// TIA Portal V21 export
FUNCTION_BLOCK "PR_5by3CylModWoRdlck"   // FB178, LAD
TITLE = 5/3Cylinder Module Without Rod Lock
{ S7_Optimized_Access := 'TRUE' }
// stored: IsIECCheckEnabled true, MemoryReserve 100, SetENOAutomatically false
   VAR_INPUT
      iResetModule : Bool;   // Reset if 1
      iResetFaults : Bool;   // Reset Fault CMD
      iEnergizeAtPwrOn : Bool;   // Energize Poweron Input
      iWorkCmd : Bool;   // Cyl Work Postion CMD
      iHomeCmd : Bool;   // Cyl Home Postion CMD
      iWorkSen : Bool;   // Cyl Work Postion Input
      iHomeSen : Bool;   // Cyl Home Postion Input
      iWorkCleartoMove : Bool;   // connect work position interlock condition healthy
      iHomeCleartoMove : Bool;   // connect home position interlock condition healthy
      iWorkPositionLeftOption : Bool;   // It is the selection of the to keep work solenoid coil on after reaching work position
      iHomePositionLeftOption : Bool;   // It is the selection of the to keep home solenoid coil on after reaching home position
      iTimeoutValue : Time;   // Time Required E.g T#500MS,T#2S
      iWorkSensDebounceVal : Time;   // Time Required E.g T#500MS,T#2S
      iHomeSensDebounceVal : Time;   // Time Required E.g T#500MS,T#2S
   END_VAR
   VAR_OUTPUT
      qWorkSol : Bool;   // Cyl Work Position Sol Output
      qHomeSol : Bool;   // Cyl Home Position Sol Output
      qWorkOver : Bool;   // 1 if Cyl at Work Position
      qHomeOver : Bool;   // 1 if Cyl at Home Position
      qModError : Bool;   // Module Error
      qErrBothSensorOn : Bool;   // 1 If both WorkSen and HomeSen inputs are high at the same time.
      qErrHomeInterlock : Bool;   // 1 If homeCleartoMove is low and home command is active.
      qErrHomeSenNotLeft : Bool;   // 1 If home position sensor did not turn off within defined time
      qErrHomeTout : Bool;   // 1 If cylinder did not reach home position within defined time
      qErrWorkInterlock : Bool;   // 1 If WorkCleartoMove is low and work command is active.
      qErrWorkSenNotLeft : Bool;   // 1 If work position sensor did not turn off within defined time
      qErrWorkTout : Bool;   // 1 If cylinder did not reach work position within defined time
      qMsgWorkPosLost : Bool;   // 1 If work position achieved and lost its position without home
      qMsgHomePosLost : Bool;   // 1 If home position achieved and lost its position without work
      qMsgBothCmdOn : Bool;   // 1 if Home & work position command on same time
   END_VAR
   VAR
      sFltRstPls : Bool;   // Stat bit for positive edge of reset fault input
      sFltEdge : Bool;   // Positive edge of fault reset input
      sWorkPosMemBit : Bool;   // Stat bit for work position memory bit
      sHomePosMemBit : Bool;   // Stat bit for Home position memory bit
      sModError : Bool;   // Stat bit for Module error
      sWorkSensDebTime : Time;   // Stat bit work sensor debounce time
      sHomeSensDebTime : Time;   // Stat bit work sensor debounce time
      sTimeoutValue : Time;   // Stat bit for time out value
      sElapsedTime : Time;   // Stat bit for time elapsed
      sDlyWorkSensDeb { S7_SetPoint := 'True'} : TON_TIME;   // On Delay for Work Sensor Debounce
      sDlyHomeSensDeb { S7_SetPoint := 'True'} : TON_TIME;   // On Delay For Home Sensor Debounce
      sDlyTimeOut { S7_SetPoint := 'True'} : TON_TIME;   // On Delay Time Out timer
      sWorkSol : Bool;
      sErrWorkTout : Bool;
      sHomeSol : Bool;
      sErrHomeTout : Bool;
      sErrBothSensorOn : Bool;
      sErrWorkInterlock : Bool;
      sErrHomeInterlock : Bool;
      sErrWorkSenNotLeft : Bool;
      sErrHomeSenNotLeft : Bool;
      sMsgHomePosLost : Bool;
      sMsgWorkPosLost : Bool;
      sPosEdge : Bool;
      sPosEdge1 : Bool;
      sRegainWrkPos : Bool;
      sRegainHomePos : Bool;
      sBothCmdOn : Bool;
      sWorkPositionLeft : Bool;
      sHomePositionLeft : Bool;
   END_VAR
   VAR_TEMP   // added for the SCL form of the ladder/FBD networks
      _w1 : Bool;
      _w2 : Bool;
      _w3 : Bool;
      _w4 : Bool;
      _w5 : Bool;
   END_VAR
BEGIN

REGION Network 1: Header
   // ==============================================================================
   //  Company: Precision Automation & Robotics India Ltd. 
   // ------------------------------------------------------------------------------
   //  Item Code:SM0101022005
   //  Author/Created by: Amiya Das
   //  Reviewed/Checked by: Atul Patwardhan
   //  First Release on: 20-01-2017
   //  Latest update on:27-01-2025 
   // ------------------------------------------------------------------------------
   //  Tested with:Simulator
   //  Engineering/Editor: TIA Portal 15 & Higher
   // ------------------------------------------------------------------------------
   //  Restrictions: No
   //  Dependencies/Requirements: NA
   // ------------------------------------------------------------------------------
   //  Change Log:
   //  Ver.	Date                            Changed by                                  Details of changes
   //  0.2           20-01-2017                  Amiya Das      	              Second release version
   //  0.3           27-01-2025                 Sujeet Rote                                qMsgBothCmdOn message is added
   //  0.4           29-01-2025                  Sujeet Rote                                Work & home position left option bit
   // ------------------------------------------------------------------------------
   // Functionality: This block is used to control a simple motion with one work 
   // position output, one home position  output, one work position sensor and one 
   // home position sensor.
   // Inputs
   // iResetModule	Bool
   // iResetFaults	Bool
   // iEnergizeAtPwrOn	Bool
   // iWorkCmd	Bool
   // iHomeCmd	Bool
   // iWorkSen	Bool
   // iHomeSen	Bool
   // iWorkCleartoMove	Bool
   // iHomeCleartoMove	Bool
   // iWorkPositionLeftOption	Bool
   // iHomePositionLeftOption	Bool
   // iTimeoutValue	Time
   // iWorkSensDebounceVal	Time
   // iHomeSensDebounceVal	Time
   // 
   // Outputs
   // qWorkSol	Bool
   // qHomeSol	Bool
   // qWorkOver	Bool
   // qHomeOver	Bool
   // qErrBothSensorOn	Bool
   // qErrHomeInterlock	Bool
   // qErrHomeSenNotLeft	Bool
   // qErrHomeTout	Bool
   // qErrWorkInterlock	Bool
   // qErrWorkSenNotLeft	Bool
   // qErrWorkTout	Bool
   // qMsgWorkPosLost	Bool
   // qMsgHomePosLost	Bool
   // qMsgBothCmdOn	Bool
   // 
   // In-outs
   // NIL
   // ------------------------------------------------------------------------------
   // Errors reported:
   // 1.qErrBothSensorOn: If both WorkSen and HomeSen inputs are high at the same time.          
   // 2.qErrHomeInterlock: If homeCleartoMove is low and home command is active.
   // 3.qErrHomeSenNotLeft: If home position sensor did not turn off within defined time 
   // 4.qErrHomeTout: If cylinder did not reach home position within defined time 
   // 5.qErrWorkInterlock: If WorkCleartoMove is low and work command is active. 
   // 7.qErrWorkSenNotLeft: If work position sensor did not turn off within defined time 
   // 8.qErrWorkTout: If cylinder did not reach work position within defined time 
   // 9.qErrPipeSwaped: If Pipe or sensor swapped
   // 
   // Messages reported:
   // 1.qMsgHomePosLost: If home position achieved and lost its position without work
   // 2.qMsgWorkPosLost: If work position achieved and lost its position without home 
   // 3.qMsgBothCmdOn :  Home & work position command on same time
   // ==============================================================================
END_REGION

REGION Network 2: Fault Reset Pulse
   // Fault Reset Pulse
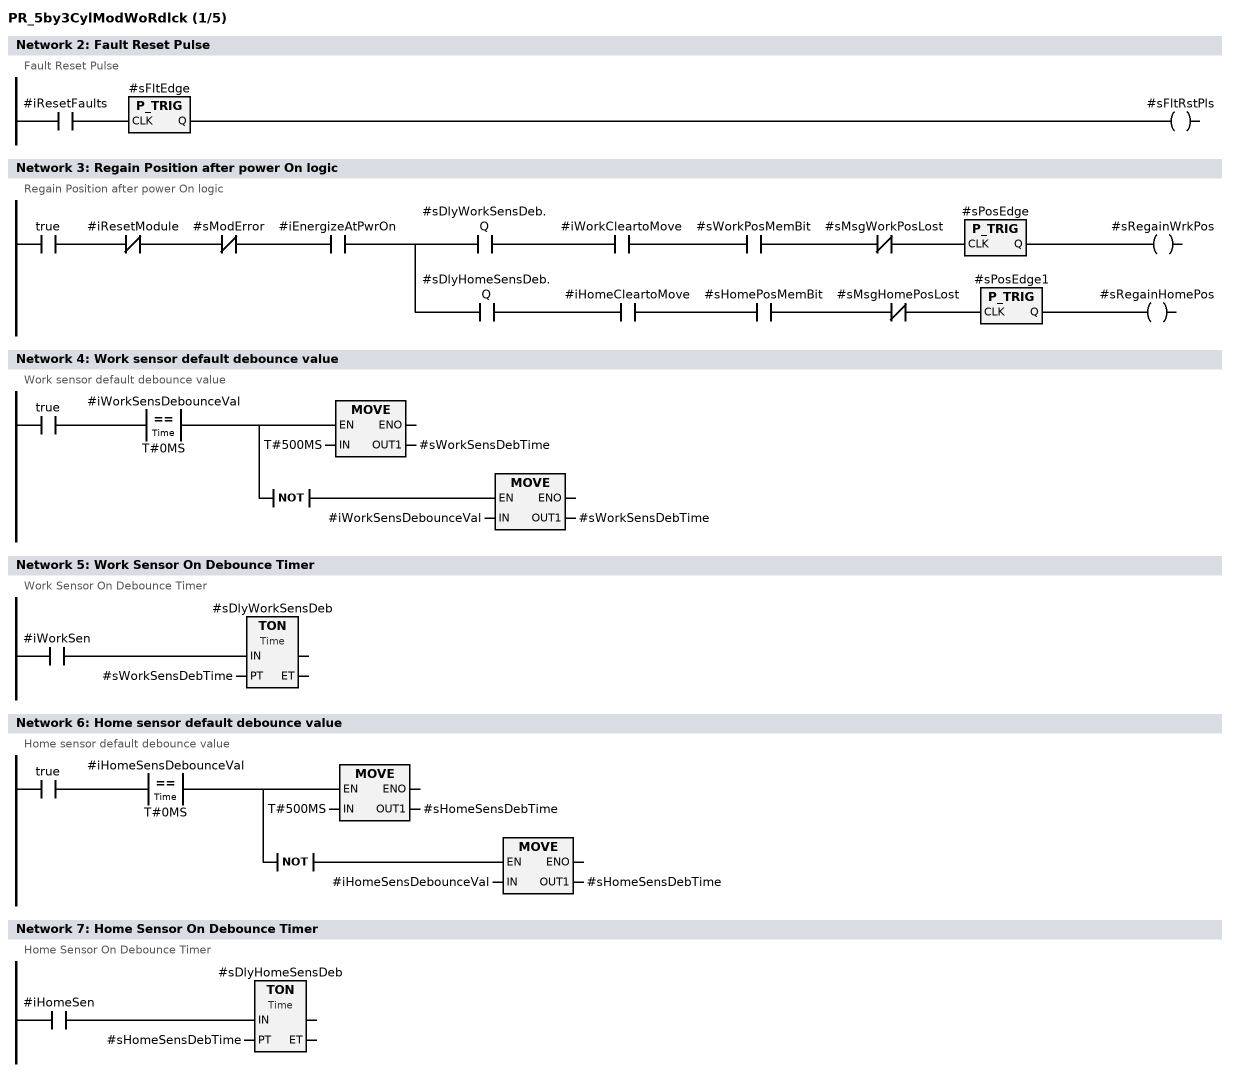
   RUNG wire#powerrail
      Contact( #iResetFaults )
      P_Trig( #sFltEdge )
      Coil( #sFltRstPls )
   END_RUNG
   // the same network as SCL:
   #_w1 := #iResetFaults AND NOT #sFltEdge;   // rising edge
   #sFltEdge := #iResetFaults;
   #sFltRstPls := #_w1;
END_REGION

REGION Network 3: Regain Position after power On logic
   // Regain Position after power On logic
   RUNG wire#powerrail
      Contact( true )
      I_Contact( #iResetModule )
      I_Contact( #sModError )
      Contact( #iEnergizeAtPwrOn )
      wire#w1
      Contact( #sDlyWorkSensDeb.Q )
      Contact( #iWorkCleartoMove )
      Contact( #sWorkPosMemBit )
      I_Contact( #sMsgWorkPosLost )
      P_Trig( #sPosEdge )
      Coil( #sRegainWrkPos )
   END_RUNG
   RUNG wire#w1
      Contact( #sDlyHomeSensDeb.Q )
      Contact( #iHomeCleartoMove )
      Contact( #sHomePosMemBit )
      I_Contact( #sMsgHomePosLost )
      P_Trig( #sPosEdge1 )
      Coil( #sRegainHomePos )
   END_RUNG
   // the same network as SCL:
   #_w1 := true AND NOT #iResetModule AND NOT #sModError AND #iEnergizeAtPwrOn;
   #_w2 := #_w1 AND #sDlyWorkSensDeb.Q AND #iWorkCleartoMove AND #sWorkPosMemBit AND NOT #sMsgWorkPosLost;
   #_w3 := #_w2 AND NOT #sPosEdge;   // rising edge
   #sPosEdge := #_w2;
   #sRegainWrkPos := #_w3;
   #_w4 := #_w1 AND #sDlyHomeSensDeb.Q AND #iHomeCleartoMove AND #sHomePosMemBit AND NOT #sMsgHomePosLost;
   #_w5 := #_w4 AND NOT #sPosEdge1;   // rising edge
   #sPosEdge1 := #_w4;
   #sRegainHomePos := #_w5;
END_REGION

REGION Network 4: Work sensor default debounce value
   // Work sensor default debounce value
   RUNG wire#powerrail
      Contact( true )
      { S7_Templates := "SrcType := Time" } EQ_Contact(in1 := #iWorkSensDebounceVal, in2 := T#0MS)
      wire#w1
      Move(in := T#500MS, out1 => #sWorkSensDebTime)
   END_RUNG
   RUNG wire#w1
      Not()
      Move(in := #iWorkSensDebounceVal, out1 => #sWorkSensDebTime)
   END_RUNG
   // the same network as SCL:
   #_w1 := true AND (#iWorkSensDebounceVal = T#0MS);
   IF #_w1 THEN #sWorkSensDebTime := T#500MS; END_IF;
   IF NOT #_w1 THEN #sWorkSensDebTime := #iWorkSensDebounceVal; END_IF;
END_REGION

REGION Network 5: Work Sensor On Debounce Timer
   // Work Sensor On Debounce Timer
   RUNG wire#powerrail
      Contact( #iWorkSen )
      { S7_Templates := "time_type := Time" } #sDlyWorkSensDeb.TON(pt := #sWorkSensDebTime, et =>)
   END_RUNG
   // the same network as SCL:
   #sDlyWorkSensDeb(IN := #iWorkSen, PT := #sWorkSensDebTime);   // TON
END_REGION

REGION Network 6: Home sensor default debounce value
   // Home sensor default debounce value
   RUNG wire#powerrail
      Contact( true )
      { S7_Templates := "SrcType := Time" } EQ_Contact(in1 := #iHomeSensDebounceVal, in2 := T#0MS)
      wire#w1
      Move(in := T#500MS, out1 => #sHomeSensDebTime)
   END_RUNG
   RUNG wire#w1
      Not()
      Move(in := #iHomeSensDebounceVal, out1 => #sHomeSensDebTime)
   END_RUNG
   // the same network as SCL:
   #_w1 := true AND (#iHomeSensDebounceVal = T#0MS);
   IF #_w1 THEN #sHomeSensDebTime := T#500MS; END_IF;
   IF NOT #_w1 THEN #sHomeSensDebTime := #iHomeSensDebounceVal; END_IF;
END_REGION

REGION Network 7: Home Sensor On Debounce Timer
   // Home Sensor On Debounce Timer
   RUNG wire#powerrail
      Contact( #iHomeSen )
      { S7_Templates := "time_type := Time" } #sDlyHomeSensDeb.TON(pt := #sHomeSensDebTime, et =>)
   END_RUNG
   // the same network as SCL:
   #sDlyHomeSensDeb(IN := #iHomeSen, PT := #sHomeSensDebTime);   // TON
END_REGION

REGION Network 8: Timeout Value
   // Timeout Value
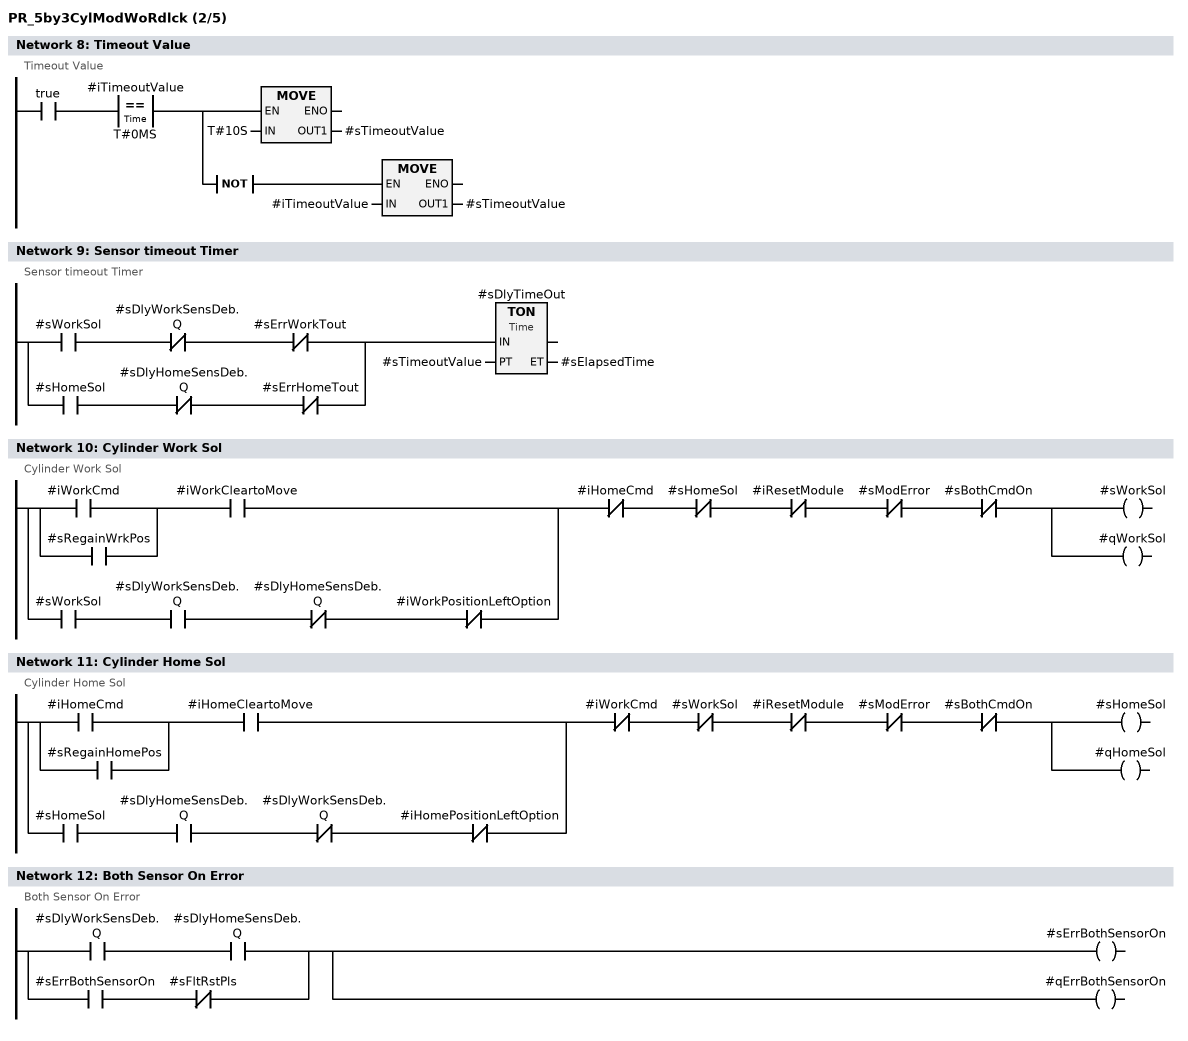
   RUNG wire#powerrail
      Contact( true )
      { S7_Templates := "SrcType := Time" } EQ_Contact(in1 := #iTimeoutValue, in2 := T#0MS)
      wire#w1
      Move(in := T#10S, out1 => #sTimeoutValue)
   END_RUNG
   RUNG wire#w1
      Not()
      Move(in := #iTimeoutValue, out1 => #sTimeoutValue)
   END_RUNG
   // the same network as SCL:
   #_w1 := true AND (#iTimeoutValue = T#0MS);
   IF #_w1 THEN #sTimeoutValue := T#10S; END_IF;
   IF NOT #_w1 THEN #sTimeoutValue := #iTimeoutValue; END_IF;
END_REGION

REGION Network 9: Sensor timeout Timer
   // Sensor timeout Timer
   RUNG wire#powerrail
      Contact( #sWorkSol )
      I_Contact( #sDlyWorkSensDeb.Q )
      I_Contact( #sErrWorkTout )
      wire#w1
      { S7_Templates := "time_type := Time" } #sDlyTimeOut.TON(pt := #sTimeoutValue, et => #sElapsedTime)
   END_RUNG
   RUNG wire#powerrail
      Contact( #sHomeSol )
      I_Contact( #sDlyHomeSensDeb.Q )
      I_Contact( #sErrHomeTout )
   END_RUNG wire#w1
   // the same network as SCL:
   #sDlyTimeOut(IN := (#sWorkSol AND NOT #sDlyWorkSensDeb.Q AND NOT #sErrWorkTout) OR (#sHomeSol AND NOT #sDlyHomeSensDeb.Q AND NOT #sErrHomeTout),   // TON
                PT := #sTimeoutValue,
                ET => #sElapsedTime);
END_REGION

REGION Network 10: Cylinder Work Sol
   // Cylinder Work Sol
   RUNG wire#powerrail
      Contact( #iWorkCmd )
      wire#w1
      Contact( #iWorkCleartoMove )
      wire#w2
      I_Contact( #iHomeCmd )
      I_Contact( #sHomeSol )
      I_Contact( #iResetModule )
      I_Contact( #sModError )
      I_Contact( #sBothCmdOn )
      wire#w3
      Coil( #sWorkSol )
   END_RUNG
   RUNG wire#powerrail
      Contact( #sRegainWrkPos )
   END_RUNG wire#w1
   RUNG wire#powerrail
      Contact( #sWorkSol )
      Contact( #sDlyWorkSensDeb.Q )
      I_Contact( #sDlyHomeSensDeb.Q )
      I_Contact( #iWorkPositionLeftOption )
   END_RUNG wire#w2
   RUNG wire#w3
      Coil( #qWorkSol )
   END_RUNG
   // the same network as SCL:
   #sWorkSol := (((#iWorkCmd OR #sRegainWrkPos) AND #iWorkCleartoMove) OR (#sWorkSol AND #sDlyWorkSensDeb.Q AND NOT #sDlyHomeSensDeb.Q AND NOT #iWorkPositionLeftOption)) AND NOT #iHomeCmd AND NOT #sHomeSol AND NOT #iResetModule AND NOT #sModError AND NOT #sBothCmdOn;
   #qWorkSol := #sWorkSol;
END_REGION

REGION Network 11: Cylinder Home Sol
   // Cylinder Home Sol
   RUNG wire#powerrail
      Contact( #iHomeCmd )
      wire#w1
      Contact( #iHomeCleartoMove )
      wire#w2
      I_Contact( #iWorkCmd )
      I_Contact( #sWorkSol )
      I_Contact( #iResetModule )
      I_Contact( #sModError )
      I_Contact( #sBothCmdOn )
      wire#w3
      Coil( #sHomeSol )
   END_RUNG
   RUNG wire#powerrail
      Contact( #sRegainHomePos )
   END_RUNG wire#w1
   RUNG wire#powerrail
      Contact( #sHomeSol )
      Contact( #sDlyHomeSensDeb.Q )
      I_Contact( #sDlyWorkSensDeb.Q )
      I_Contact( #iHomePositionLeftOption )
   END_RUNG wire#w2
   RUNG wire#w3
      Coil( #qHomeSol )
   END_RUNG
   // the same network as SCL:
   #sHomeSol := (((#iHomeCmd OR #sRegainHomePos) AND #iHomeCleartoMove) OR (#sHomeSol AND #sDlyHomeSensDeb.Q AND NOT #sDlyWorkSensDeb.Q AND NOT #iHomePositionLeftOption)) AND NOT #iWorkCmd AND NOT #sWorkSol AND NOT #iResetModule AND NOT #sModError AND NOT #sBothCmdOn;
   #qHomeSol := #sHomeSol;
END_REGION

REGION Network 12: Both Sensor On Error
   // Both Sensor On Error
   RUNG wire#powerrail
      Contact( #sDlyWorkSensDeb.Q )
      Contact( #sDlyHomeSensDeb.Q )
      wire#w1
      Coil( #sErrBothSensorOn )
   END_RUNG
   RUNG wire#powerrail
      Contact( #sErrBothSensorOn )
      I_Contact( #sFltRstPls )
   END_RUNG wire#w1
   RUNG wire#w1
      Coil( #qErrBothSensorOn )
   END_RUNG
   // the same network as SCL:
   #sErrBothSensorOn := (#sDlyWorkSensDeb.Q AND #sDlyHomeSensDeb.Q) OR (#sErrBothSensorOn AND NOT #sFltRstPls);
   #qErrBothSensorOn := #sErrBothSensorOn;
END_REGION

REGION Network 13: Work Interlock Error
   // Work Interlock Error
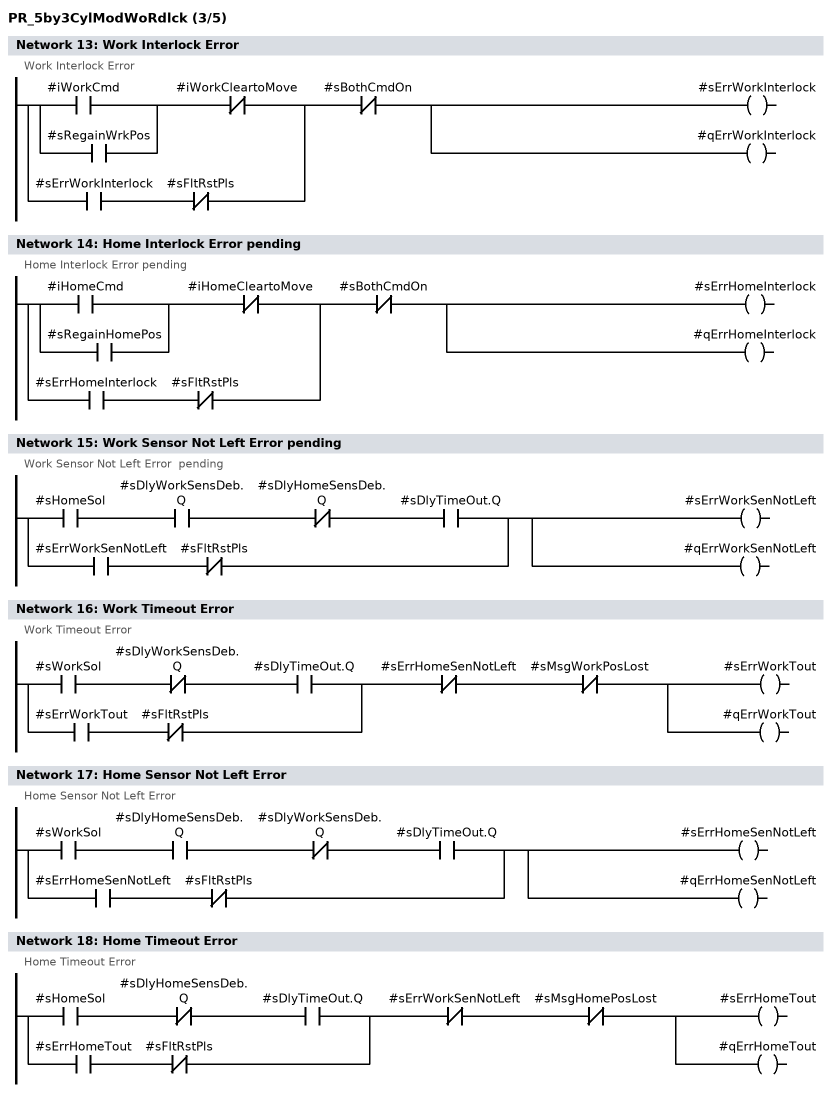
   RUNG wire#powerrail
      Contact( #iWorkCmd )
      wire#w1
      I_Contact( #iWorkCleartoMove )
      wire#w2
      I_Contact( #sBothCmdOn )
      wire#w3
      Coil( #sErrWorkInterlock )
   END_RUNG
   RUNG wire#powerrail
      Contact( #sRegainWrkPos )
   END_RUNG wire#w1
   RUNG wire#powerrail
      Contact( #sErrWorkInterlock )
      I_Contact( #sFltRstPls )
   END_RUNG wire#w2
   RUNG wire#w3
      Coil( #qErrWorkInterlock )
   END_RUNG
   // the same network as SCL:
   #sErrWorkInterlock := (((#iWorkCmd OR #sRegainWrkPos) AND NOT #iWorkCleartoMove) OR (#sErrWorkInterlock AND NOT #sFltRstPls)) AND NOT #sBothCmdOn;
   #qErrWorkInterlock := #sErrWorkInterlock;
END_REGION

REGION Network 14: Home Interlock Error pending
   // Home Interlock Error pending
   RUNG wire#powerrail
      Contact( #iHomeCmd )
      wire#w1
      I_Contact( #iHomeCleartoMove )
      wire#w2
      I_Contact( #sBothCmdOn )
      wire#w3
      Coil( #sErrHomeInterlock )
   END_RUNG
   RUNG wire#powerrail
      Contact( #sRegainHomePos )
   END_RUNG wire#w1
   RUNG wire#powerrail
      Contact( #sErrHomeInterlock )
      I_Contact( #sFltRstPls )
   END_RUNG wire#w2
   RUNG wire#w3
      Coil( #qErrHomeInterlock )
   END_RUNG
   // the same network as SCL:
   #sErrHomeInterlock := (((#iHomeCmd OR #sRegainHomePos) AND NOT #iHomeCleartoMove) OR (#sErrHomeInterlock AND NOT #sFltRstPls)) AND NOT #sBothCmdOn;
   #qErrHomeInterlock := #sErrHomeInterlock;
END_REGION

REGION Network 15: Work Sensor Not Left Error pending
   // Work Sensor Not Left Error  pending
   RUNG wire#powerrail
      Contact( #sHomeSol )
      Contact( #sDlyWorkSensDeb.Q )
      I_Contact( #sDlyHomeSensDeb.Q )
      Contact( #sDlyTimeOut.Q )
      wire#w1
      Coil( #sErrWorkSenNotLeft )
   END_RUNG
   RUNG wire#powerrail
      Contact( #sErrWorkSenNotLeft )
      I_Contact( #sFltRstPls )
   END_RUNG wire#w1
   RUNG wire#w1
      Coil( #qErrWorkSenNotLeft )
   END_RUNG
   // the same network as SCL:
   #sErrWorkSenNotLeft := (#sHomeSol AND #sDlyWorkSensDeb.Q AND NOT #sDlyHomeSensDeb.Q AND #sDlyTimeOut.Q) OR (#sErrWorkSenNotLeft AND NOT #sFltRstPls);
   #qErrWorkSenNotLeft := #sErrWorkSenNotLeft;
END_REGION

REGION Network 16: Work Timeout Error
   // Work Timeout Error
   RUNG wire#powerrail
      Contact( #sWorkSol )
      I_Contact( #sDlyWorkSensDeb.Q )
      Contact( #sDlyTimeOut.Q )
      wire#w1
      I_Contact( #sErrHomeSenNotLeft )
      I_Contact( #sMsgWorkPosLost )
      wire#w2
      Coil( #sErrWorkTout )
   END_RUNG
   RUNG wire#powerrail
      Contact( #sErrWorkTout )
      I_Contact( #sFltRstPls )
   END_RUNG wire#w1
   RUNG wire#w2
      Coil( #qErrWorkTout )
   END_RUNG
   // the same network as SCL:
   #sErrWorkTout := ((#sWorkSol AND NOT #sDlyWorkSensDeb.Q AND #sDlyTimeOut.Q) OR (#sErrWorkTout AND NOT #sFltRstPls)) AND NOT #sErrHomeSenNotLeft AND NOT #sMsgWorkPosLost;
   #qErrWorkTout := #sErrWorkTout;
END_REGION

REGION Network 17: Home Sensor Not Left Error
   // Home Sensor Not Left Error
   RUNG wire#powerrail
      Contact( #sWorkSol )
      Contact( #sDlyHomeSensDeb.Q )
      I_Contact( #sDlyWorkSensDeb.Q )
      Contact( #sDlyTimeOut.Q )
      wire#w1
      Coil( #sErrHomeSenNotLeft )
   END_RUNG
   RUNG wire#powerrail
      Contact( #sErrHomeSenNotLeft )
      I_Contact( #sFltRstPls )
   END_RUNG wire#w1
   RUNG wire#w1
      Coil( #qErrHomeSenNotLeft )
   END_RUNG
   // the same network as SCL:
   #sErrHomeSenNotLeft := (#sWorkSol AND #sDlyHomeSensDeb.Q AND NOT #sDlyWorkSensDeb.Q AND #sDlyTimeOut.Q) OR (#sErrHomeSenNotLeft AND NOT #sFltRstPls);
   #qErrHomeSenNotLeft := #sErrHomeSenNotLeft;
END_REGION

REGION Network 18: Home Timeout Error
   // Home Timeout Error
   RUNG wire#powerrail
      Contact( #sHomeSol )
      I_Contact( #sDlyHomeSensDeb.Q )
      Contact( #sDlyTimeOut.Q )
      wire#w1
      I_Contact( #sErrWorkSenNotLeft )
      I_Contact( #sMsgHomePosLost )
      wire#w2
      Coil( #sErrHomeTout )
   END_RUNG
   RUNG wire#powerrail
      Contact( #sErrHomeTout )
      I_Contact( #sFltRstPls )
   END_RUNG wire#w1
   RUNG wire#w2
      Coil( #qErrHomeTout )
   END_RUNG
   // the same network as SCL:
   #sErrHomeTout := ((#sHomeSol AND NOT #sDlyHomeSensDeb.Q AND #sDlyTimeOut.Q) OR (#sErrHomeTout AND NOT #sFltRstPls)) AND NOT #sErrWorkSenNotLeft AND NOT #sMsgHomePosLost;
   #qErrHomeTout := #sErrHomeTout;
END_REGION

REGION Network 19: Work Position Left Stat logic / Work Position Left option bit Logic
   // Work Position Left Stat logic / Work Position Left option bit Logic
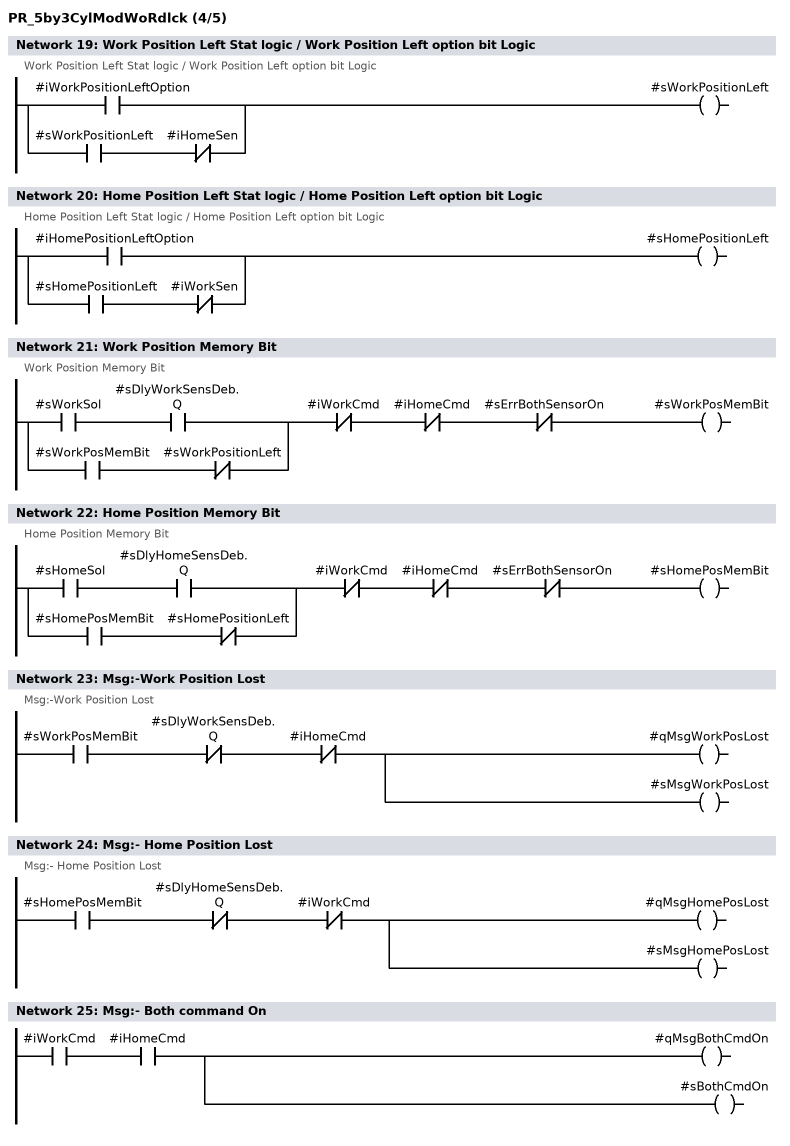
   RUNG wire#powerrail
      Contact( #iWorkPositionLeftOption )
      wire#w1
      Coil( #sWorkPositionLeft )
   END_RUNG
   RUNG wire#powerrail
      Contact( #sWorkPositionLeft )
      I_Contact( #iHomeSen )
   END_RUNG wire#w1
   // the same network as SCL:
   #sWorkPositionLeft := #iWorkPositionLeftOption OR (#sWorkPositionLeft AND NOT #iHomeSen);
END_REGION

REGION Network 20: Home Position Left Stat logic / Home Position Left option bit Logic
   // Home Position Left Stat logic / Home Position Left option bit Logic
   RUNG wire#powerrail
      Contact( #iHomePositionLeftOption )
      wire#w1
      Coil( #sHomePositionLeft )
   END_RUNG
   RUNG wire#powerrail
      Contact( #sHomePositionLeft )
      I_Contact( #iWorkSen )
   END_RUNG wire#w1
   // the same network as SCL:
   #sHomePositionLeft := #iHomePositionLeftOption OR (#sHomePositionLeft AND NOT #iWorkSen);
END_REGION

REGION Network 21: Work Position Memory Bit
   // Work Position Memory Bit
   RUNG wire#powerrail
      Contact( #sWorkSol )
      Contact( #sDlyWorkSensDeb.Q )
      wire#w1
      I_Contact( #iWorkCmd )
      I_Contact( #iHomeCmd )
      I_Contact( #sErrBothSensorOn )
      Coil( #sWorkPosMemBit )
   END_RUNG
   RUNG wire#powerrail
      Contact( #sWorkPosMemBit )
      I_Contact( #sWorkPositionLeft )
   END_RUNG wire#w1
   // the same network as SCL:
   #sWorkPosMemBit := ((#sWorkSol AND #sDlyWorkSensDeb.Q) OR (#sWorkPosMemBit AND NOT #sWorkPositionLeft)) AND NOT #iWorkCmd AND NOT #iHomeCmd AND NOT #sErrBothSensorOn;
END_REGION

REGION Network 22: Home Position Memory Bit
   // Home Position Memory Bit
   RUNG wire#powerrail
      Contact( #sHomeSol )
      Contact( #sDlyHomeSensDeb.Q )
      wire#w1
      I_Contact( #iWorkCmd )
      I_Contact( #iHomeCmd )
      I_Contact( #sErrBothSensorOn )
      Coil( #sHomePosMemBit )
   END_RUNG
   RUNG wire#powerrail
      Contact( #sHomePosMemBit )
      I_Contact( #sHomePositionLeft )
   END_RUNG wire#w1
   // the same network as SCL:
   #sHomePosMemBit := ((#sHomeSol AND #sDlyHomeSensDeb.Q) OR (#sHomePosMemBit AND NOT #sHomePositionLeft)) AND NOT #iWorkCmd AND NOT #iHomeCmd AND NOT #sErrBothSensorOn;
END_REGION

REGION Network 23: Msg:-Work Position Lost
   // Msg:-Work Position Lost
   RUNG wire#powerrail
      Contact( #sWorkPosMemBit )
      I_Contact( #sDlyWorkSensDeb.Q )
      I_Contact( #iHomeCmd )
      wire#w1
      Coil( #qMsgWorkPosLost )
   END_RUNG
   RUNG wire#w1
      Coil( #sMsgWorkPosLost )
   END_RUNG
   // the same network as SCL:
   #qMsgWorkPosLost := #sWorkPosMemBit AND NOT #sDlyWorkSensDeb.Q AND NOT #iHomeCmd;
   #sMsgWorkPosLost := #qMsgWorkPosLost;
END_REGION

REGION Network 24: Msg:- Home Position Lost
   // Msg:- Home Position Lost
   RUNG wire#powerrail
      Contact( #sHomePosMemBit )
      I_Contact( #sDlyHomeSensDeb.Q )
      I_Contact( #iWorkCmd )
      wire#w1
      Coil( #qMsgHomePosLost )
   END_RUNG
   RUNG wire#w1
      Coil( #sMsgHomePosLost )
   END_RUNG
   // the same network as SCL:
   #qMsgHomePosLost := #sHomePosMemBit AND NOT #sDlyHomeSensDeb.Q AND NOT #iWorkCmd;
   #sMsgHomePosLost := #qMsgHomePosLost;
END_REGION

REGION Network 25: Msg:- Both command On
   RUNG wire#powerrail
      Contact( #iWorkCmd )
      Contact( #iHomeCmd )
      wire#w1
      Coil( #qMsgBothCmdOn )
   END_RUNG
   RUNG wire#w1
      Coil( #sBothCmdOn )
   END_RUNG
   // the same network as SCL:
   #qMsgBothCmdOn := #iWorkCmd AND #iHomeCmd;
   #sBothCmdOn := #qMsgBothCmdOn;
END_REGION

REGION Network 26: Module Error
   // Module Error
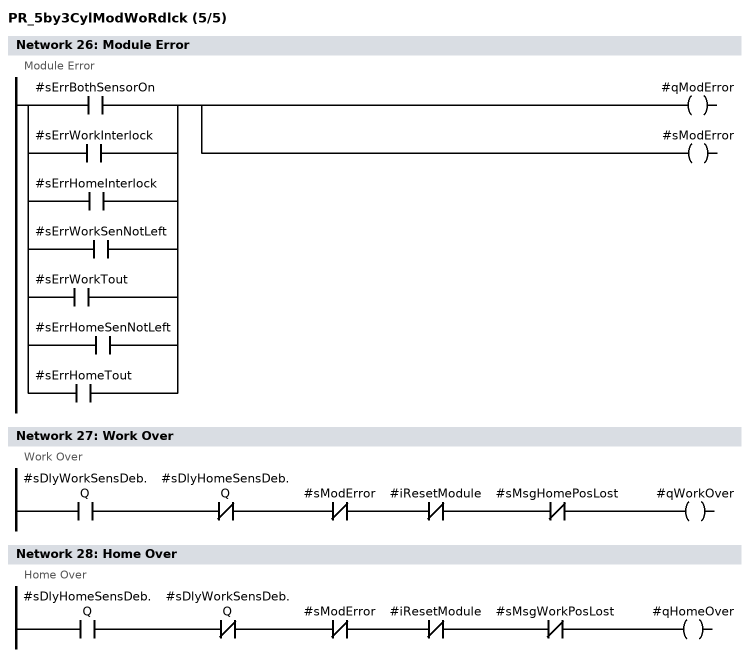
   RUNG wire#powerrail
      Contact( #sErrBothSensorOn )
      wire#w1
      Coil( #qModError )
   END_RUNG
   RUNG wire#powerrail
      Contact( #sErrWorkInterlock )
   END_RUNG wire#w1
   RUNG wire#powerrail
      Contact( #sErrHomeInterlock )
   END_RUNG wire#w1
   RUNG wire#powerrail
      Contact( #sErrWorkSenNotLeft )
   END_RUNG wire#w1
   RUNG wire#powerrail
      Contact( #sErrWorkTout )
   END_RUNG wire#w1
   RUNG wire#powerrail
      Contact( #sErrHomeSenNotLeft )
   END_RUNG wire#w1
   RUNG wire#powerrail
      Contact( #sErrHomeTout )
   END_RUNG wire#w1
   RUNG wire#w1
      Coil( #sModError )
   END_RUNG
   // the same network as SCL:
   #qModError := #sErrBothSensorOn OR #sErrWorkInterlock OR #sErrHomeInterlock OR #sErrWorkSenNotLeft OR #sErrWorkTout OR #sErrHomeSenNotLeft OR #sErrHomeTout;
   #sModError := #qModError;
END_REGION

REGION Network 27: Work Over
   // Work Over
   RUNG wire#powerrail
      Contact( #sDlyWorkSensDeb.Q )
      I_Contact( #sDlyHomeSensDeb.Q )
      I_Contact( #sModError )
      I_Contact( #iResetModule )
      I_Contact( #sMsgHomePosLost )
      Coil( #qWorkOver )
   END_RUNG
   // the same network as SCL:
   #qWorkOver := #sDlyWorkSensDeb.Q AND NOT #sDlyHomeSensDeb.Q AND NOT #sModError AND NOT #iResetModule AND NOT #sMsgHomePosLost;
END_REGION

REGION Network 28: Home Over
   // Home Over
   RUNG wire#powerrail
      Contact( #sDlyHomeSensDeb.Q )
      I_Contact( #sDlyWorkSensDeb.Q )
      I_Contact( #sModError )
      I_Contact( #iResetModule )
      I_Contact( #sMsgWorkPosLost )
      Coil( #qHomeOver )
   END_RUNG
   // the same network as SCL:
   #qHomeOver := #sDlyHomeSensDeb.Q AND NOT #sDlyWorkSensDeb.Q AND NOT #sModError AND NOT #iResetModule AND NOT #sMsgWorkPosLost;
END_REGION
END_FUNCTION_BLOCK
